Staubli VAL3: selMainProg.pgx

public program selMainProg()
begin
  nProgType=2
end
